FUNCTION_BLOCK F (* Positive: shared prelude holding a lowered timer, whose X_STATE beside X_START_TIME is not a control position *)
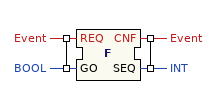
  EVENT_INPUT
    REQ WITH GO;
  END_EVENT
  EVENT_OUTPUT
    CNF WITH SEQ;
  END_EVENT
  VAR_INPUT
    GO : BOOL;
  END_VAR
  VAR_OUTPUT
    SEQ : INT;
  END_VAR
  VAR
    T_STATE : INT;
    T_PREV_IN : BOOL;
    T_Q : BOOL;
    T_START_TIME : TIME;
    NOW : TIME;
  END_VAR
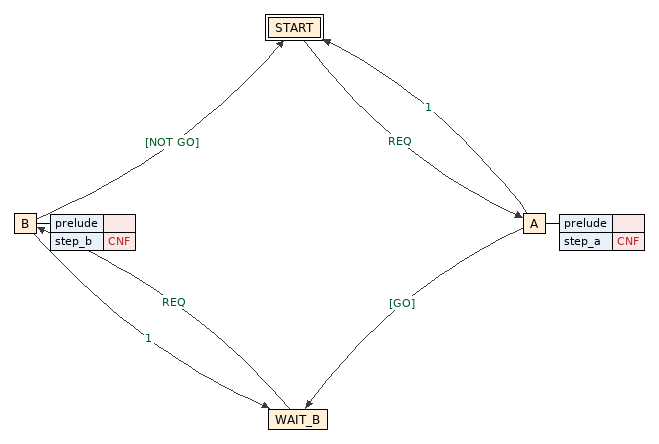
  EC_STATES
    START;
    A : prelude, step_a -> CNF;
    WAIT_B;
    B : prelude, step_b -> CNF;
  END_STATES
  EC_TRANSITIONS
    START TO A := REQ;
    A TO WAIT_B := [GO];
    A TO START := 1;
    WAIT_B TO B := REQ;
    B TO START := [NOT GO];
    B TO WAIT_B := 1;
  END_TRANSITIONS
  ALGORITHM prelude IN ST:
NOW := NOW + T#10ms;
IF (T_STATE = 0) AND NOT T_PREV_IN AND GO THEN
  T_STATE := 1;
  T_Q := FALSE;
  T_START_TIME := NOW;
ELSE
  IF NOT GO THEN
    T_Q := FALSE;
    T_STATE := 0;
  ELSIF T_STATE = 1 THEN
    IF T_START_TIME + T#50ms <= NOW THEN
      T_STATE := 2;
      T_Q := TRUE;
    END_IF;
  END_IF;
END_IF;
T_PREV_IN := GO;
  END_ALGORITHM
  ALGORITHM step_a IN ST:
SEQ := 0;
IF GO THEN
  SEQ := 1;
END_IF;
  END_ALGORITHM
  ALGORITHM step_b IN ST:
IF NOT GO THEN
  SEQ := 0;
END_IF;
  END_ALGORITHM
END_FUNCTION_BLOCK
